ABB RobotStudio station: Caja2Inclinada.rspag

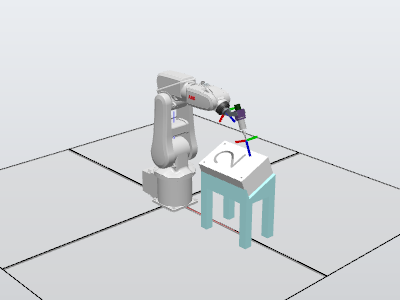
--- station ---
Station Project6 (saved by RobotStudio 26.3.11794.0)
Controller IRB120_3_58
  mechanical unit ROB_1: IRB120_3_58__01, 6 joints, base frame (0, 0, 0) mm
Layout (positions relative to the parent item):
  - IRB120_3_58__01 [mechanism, from %ABB.RobotStudio.Models.IRB120%\IRB120_3_58_G_01.rslib] at (0, 0, 0) mm; joint values [0, 0, 0, 0, 0.5236, 0] (rad or m)
  - punta [mechanism, from Components\punta.rslib] at (364.35, 0, 594) mm, rotated rx 180 ry 60 rz 180 deg
  - CajaNumero2 [part] at (585.43, -73.22, 252.41) mm, rotated rx 0 ry -22.39 rz 90.07 deg, size 188.7 x 287.5 x 103.3 mm
  - mesarRobotStudio [part] at (600, 98.92, 2.52) mm, rotated rx 0.01 ry 0 rz -179.93 deg, size 304.8 x 198.1 x 325.1 mm
Attachment: punta is attached to IRB120_3_58__01 / Link6
Collision set Conjunto de colisión_1: CajaNumero2 against punta, near miss 0 m
Targets, tools, work objects and paths stored in the station and not in the controller backup, written as RAPID:
! task T_ROB1
MODULE CalibData
  PERS tooldata punta:=[TRUE,[[24,0,172],[0.945518576,0,0.325568154,0]],[0.1,[0,0,1],[1,0,0,0],0,0,0]];
ENDMODULE


--- Controller Data/IRB120_3_58/RAPID/TASK1/PROGMOD/Module1.mod ---
MODULE Module1
    !***********************************************************
    !
    ! M?dulo:  Module1
    !
    ! Descripción:
    !   <Introduzca la descripción aquí>
    !
    ! Autor: ferna
    !
    ! Versión: 1.0
    !
    !***********************************************************


    !***********************************************************
    !
    ! Procedimiento Main
    !
    !   Este es el punto de entrada de su programa
    !
    !***********************************************************
    PROC main()
        !Add your code here
    ENDPROC
ENDMODULE
